(*
SPDX-FileCopyrightText: © 2026 Oleksandr Tiutyk <trofimich@gmail.com>
SPDX-License-Identifier: MIT
License: https://opensource.org/license/mit
*)

(*!
<summary>Marker interface representing an embedded condition reset scope node.</summary>
<description>
Scopes are linked in an ownership tree to restore variable state during condition resets.
Instances are non-copyable, owned by an activity or condition, and managed within a single task.
</description>
*)
{attribute 'hide'}
INTERFACE IVariableResetScope EXTENDS TOF_Core.IObject

END_INTERFACE

(* stored: Version 1.1.0.1
   Itf IVariableResetScope: Id {4e5ac262-ddbc-45f3-a2c6-572ffed731fb} *)
